% RSLogix 500 project packaging machine.RSS, saved by version 8.30.00.16 %
PROJECT "UNTITLED"    % processor: MicroLogix 1000 %

PROGRAM FILES
  LAD 2 "MAIN_PROG"  8 rungs
  LAD 3 "USER_FAULT"  1 rungs
  LAD 4 "HSC_INT"  1 rungs
  LAD 5 "STI_INT"  1 rungs
  LAD 6, 7, 8, 9, 10, 11, 12, 13, 14, 15, 16: only END

DATA FILES
  O0 OUTPUT  5 elements
  I1 INPUT  8 elements
  S2 STATUS  33 elements
  B3 BINARY  32 elements
  T4 TIMER  40 elements
  C5 COUNTER  32 elements
  R6 CONTROL  16 elements
  N7 INTEGER  105 elements

LADDER 2 "MAIN_PROG"
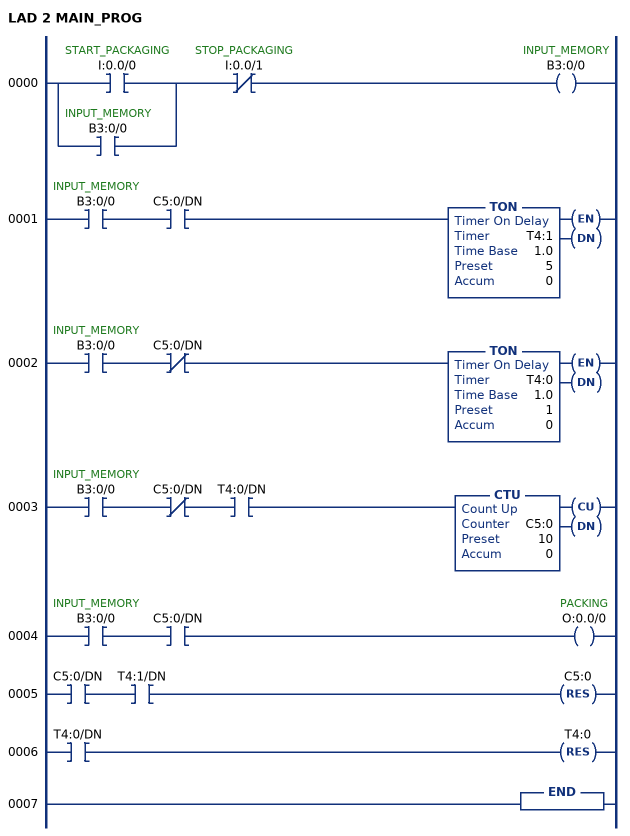
% Rung: 0 %
SOR BST XIC I:0.0/0 NXB XIC B3:0/0 BND XIO I:0.0/1 OTE B3:0/0 EOR
%   I:0.0/0  START_PACKAGING %
%   B3:0/0  INPUT_MEMORY %
%   I:0.0/1  STOP_PACKAGING %
% Rung: 1 %
SOR XIC B3:0/0 XIC C5:0/DN TON T4:1 1.0 5 0 EOR
%   B3:0/0  INPUT_MEMORY %
% Rung: 2 %
SOR XIC B3:0/0 XIO C5:0/DN TON T4:0 1.0 1 0 EOR
%   B3:0/0  INPUT_MEMORY %
% Rung: 3 %
SOR XIC B3:0/0 XIO C5:0/DN XIC T4:0/DN CTU C5:0 10 0 EOR
%   B3:0/0  INPUT_MEMORY %
% Rung: 4 %
SOR XIC B3:0/0 XIC C5:0/DN OTE O:0.0/0 EOR
%   B3:0/0  INPUT_MEMORY %
%   O:0.0/0  PACKING %
% Rung: 5 %
SOR XIC C5:0/DN XIC T4:1/DN RES C5:0 EOR
% Rung: 6 %
SOR XIC T4:0/DN RES T4:0 EOR
% Rung: 7 %
SOR END EOR

DATA TABLE (non-zero values as saved)
DATA T4
% .PRE .ACC %
% T4:0 % 1 0
% T4:1 % 5 0
DATA C5
% .PRE .ACC %
% C5:0 % 10 0
